{region 'Documentation'}
(*!
<summary>Checks two-sample qualification and PLC-owned clearing for one external lifecycle command.</summary>
<description>
Use one instance per Start, Abort and Reset. Every enabled cycle samples the real adapter once.
The script first withdraws two separate one-sample pulses, then leaves TRUE untouched for two
calls. Acceptance must forward exactly one request and clear that field. A following call
without a write must not repeat it. A new TRUE then needs two new samples before request two.
Each sample checks the selected count/bit and both unrelated commands. This is deterministic
call-boundary evidence, not a simulation of asynchronous ADS writes or a command handshake.
ProcessReset initializes the local subject and clears the recorder for repeatable runs.
</description>
*)
{endregion}
FUNCTION_BLOCK Test_CommandQualification EXTENDS TestCaseBase
VAR_INPUT
    Command : E_AdapterCommand := E_AdapterCommand.Start; //! External command field exercised by this instance; held fixed by the containing Suite.
END_VAR
VAR
    FSubject : RunControlCommandAdapter;
    FOwner : RunControlRequestRecorder;
    FControl : ST_RunControl;
    FStep : UINT;
    FSampleChecked : BOOL;
    FRequestCount : AssertTrue;
    FRequestCountMatches : BOOL;
    FCommandValue : AssertTrue;
    FCommandValueMatches : BOOL;
    FOtherCommands : AssertTrue;
    FOtherCommandsMatches : BOOL;
END_VAR
VAR CONSTANT
    Baseline : UINT := 0;
    SinglePulse : UINT := 1;
    Withdrawal : UINT := 2;
    SeparatedPulse : UINT := 3;
    SecondWithdrawal : UINT := 4;
    RetainedFirstSample : UINT := 5;
    RetainedSecondSample : UINT := 6;
    FreshFirstSample : UINT := 8;
    FreshSecondSample : UINT := 9;
    AfterFreshClearing : UINT := 10;
END_VAR

SUPER^();

{region 'Documentation'}
(*!
<summary>Collects request-count, field-value and isolation checks.</summary>
*)
{endregion}
METHOD PROTECTED AggregateResults
VAR_INPUT
    Aggregator : I_ResultAggregator; //! Borrowed result sink owned by the outer Test Case; add this test's checking Assertions without resetting or retaining the sink.
END_VAR
Aggregator.AddProvider(Provider := FRequestCount);
Aggregator.AddProvider(Provider := FCommandValue);
Aggregator.AddProvider(Provider := FOtherCommands);
END_METHOD

{region 'Documentation'}
(*!
<summary>Checks the explicit script oracle against recorded calls and the post-call command fields.</summary>
*)
{endregion}
METHOD PRIVATE CheckSample
VAR
    ExpectedCount : UINT;
    ExpectedCommand : BOOL;
    ActualCount : UINT;
    ActualCommand : BOOL;
END_VAR
IF FStep >= FreshSecondSample THEN
    ExpectedCount := 2;
ELSIF FStep >= RetainedSecondSample THEN
    ExpectedCount := 1;
END_IF;
ExpectedCommand := (FStep = SinglePulse) OR (FStep = SeparatedPulse)
    OR (FStep = RetainedFirstSample) OR (FStep = FreshFirstSample);
CASE Command OF
    E_AdapterCommand.Start:
        ActualCount := FOwner.StartCount;
        ActualCommand := FControl.Cmd.Start;
        FOtherCommandsMatches := (FOwner.AbortCount = 0) AND (FOwner.ResetCount = 0)
            AND NOT FControl.Cmd.Abort AND NOT FControl.Cmd.Reset;
    E_AdapterCommand.Abort:
        ActualCount := FOwner.AbortCount;
        ActualCommand := FControl.Cmd.Abort;
        FOtherCommandsMatches := (FOwner.StartCount = 0) AND (FOwner.ResetCount = 0)
            AND NOT FControl.Cmd.Start AND NOT FControl.Cmd.Reset;
    E_AdapterCommand.Reset:
        ActualCount := FOwner.ResetCount;
        ActualCommand := FControl.Cmd.Reset;
        FOtherCommandsMatches := (FOwner.StartCount = 0) AND (FOwner.AbortCount = 0)
            AND NOT FControl.Cmd.Start AND NOT FControl.Cmd.Abort;
END_CASE;
FRequestCountMatches := ActualCount = ExpectedCount;
FCommandValueMatches := ActualCommand = ExpectedCommand;
END_METHOD

{region 'Documentation'}
(*!
<summary>Initializes the three checking Assertions for the selected command.</summary>
*)
{endregion}
METHOD PROTECTED Configure
FPreparationStateCount := 0;
FTestStateCount := 1;
FRequestCount.Initialize(Parent := THIS^,
    AssertionName := 'RequestCount');
FCommandValue.Initialize(Parent := THIS^,
    AssertionName := 'CommandValue');
FOtherCommands.Initialize(Parent := THIS^,
    AssertionName := 'OtherCommands');
END_METHOD

{region 'Documentation'}
(*!
<summary>No asynchronous resource needs abort handling.</summary>
*)
{endregion}
METHOD PROTECTED ProcessAbort
VAR_INPUT
    Enable : BOOL; //! Phase permission supplied by the owning Test Case; FALSE does not authorize progression, while observation may continue.
END_VAR
IF Enable THEN
    CompleteAbort();
END_IF;
END_METHOD

{region 'Documentation'}
(*!
<summary>Checks every sample before advancing; failures remain latched across the script.</summary>
*)
{endregion}
METHOD PROTECTED ProcessAssertions
VAR_INPUT
    Enable : BOOL; //! Phase permission supplied by the owning Test Case; FALSE does not authorize progression, while observation may continue.
END_VAR
FRequestCount(Enable := Enable,
    State := State,
    IN := FRequestCountMatches);
FCommandValue(Enable := Enable,
    State := State,
    IN := FCommandValueMatches);
FOtherCommands(Enable := Enable,
    State := State,
    IN := FOtherCommandsMatches);
IF Enable THEN
    FSampleChecked := TRUE;
END_IF;
END_METHOD

{region 'Documentation'}
(*!
<summary>No Preparation work is required.</summary>
*)
{endregion}
METHOD PROTECTED ProcessPreparations
VAR_INPUT
    // SA0033: Required override; this test has no Preparation phase.
    {attribute 'analysis' := '-33'}
    Enable : BOOL; //! Phase permission supplied by the owning Test Case; FALSE does not authorize progression, while observation may continue.
END_VAR
END_METHOD

{region 'Documentation'}
(*!
<summary>Clears subject history, recorded requests and the bounded sample script.</summary>
*)
{endregion}
METHOD PROTECTED ProcessReset
FSubject.Initialize(ControlData := FControl);
FOwner.Clear();
FStep := Baseline;
FSampleChecked := FALSE;
FRequestCount.Reset();
FRequestCountMatches := FALSE;
FCommandValue.Reset();
FCommandValueMatches := FALSE;
FOtherCommands.Reset();
FOtherCommandsMatches := FALSE;
CompleteReset();
END_METHOD

{region 'Documentation'}
(*!
<summary>Applies one scheduled write and one real adapter call per active PLC cycle.</summary>
*)
{endregion}
METHOD PROTECTED ProcessTests
VAR_INPUT
    Enable : BOOL; //! Phase permission supplied by the owning Test Case; FALSE does not authorize progression, while observation may continue.
END_VAR
IF NOT Enable THEN
    RETURN;
END_IF;
IF FSampleChecked THEN
    IF FStep = AfterFreshClearing THEN
        CompleteTests();
        RETURN;
    END_IF;
    FStep := FStep + 1;
    FSampleChecked := FALSE;
END_IF;
CASE FStep OF
    SinglePulse, SeparatedPulse, RetainedFirstSample, FreshFirstSample:
        SetCommand(Value := TRUE);
    Withdrawal, SecondWithdrawal:
        SetCommand(Value := FALSE);
ELSE
    // No external write: retain the actual field, including the adapter's clearing.
END_CASE;
FSubject(RunControl := FOwner,
    Commands := FControl.Cmd);
CheckSample();
END_METHOD

{region 'Documentation'}
(*!
<summary>Writes only the chosen external command field.</summary>
*)
{endregion}
METHOD PRIVATE SetCommand
VAR_INPUT
    Value : BOOL; //! Boolean value written only to the selected command field.
END_VAR
CASE Command OF
    E_AdapterCommand.Start:
        FControl.Cmd.Start := Value;
    E_AdapterCommand.Abort:
        FControl.Cmd.Abort := Value;
    E_AdapterCommand.Reset:
        FControl.Cmd.Reset := Value;
END_CASE;
END_METHOD

END_FUNCTION_BLOCK

(* stored: Version 1.1.0.1
   POU Test_CommandQualification: Id {4653a244-9dde-40c4-bba8-7d26f3686632}, SpecialFunc None
   Folder Internal: Id {49490200-0000-4000-8000-000000000001}
   Method AggregateResults: Id {49490200-0000-4000-8000-000000000003}
   Method CheckSample: Id {49490200-0000-4000-8000-000000000008}
   Method Configure: Id {49490200-0000-4000-8000-000000000002}
   Method ProcessAbort: Id {49490200-0000-4000-8000-000000000005}
   Method ProcessAssertions: Id {49490200-0000-4000-8000-000000000010}
   Method ProcessPreparations: Id {49490200-0000-4000-8000-000000000006}
   Method ProcessReset: Id {49490200-0000-4000-8000-000000000004}
   Method ProcessTests: Id {49490200-0000-4000-8000-000000000009}
   Method SetCommand: Id {49490200-0000-4000-8000-000000000007} *)
